// TIA Portal V20 export
// export: Created 2026-10-19T18:06:23.6211165Z, ExportSetting WithDefaults, DisplayName Totally Integrated Automation Portal, DisplayVersion V20 Update 6, DisplayName TIA Portal Openness, DisplayVersion V20 Update 6, DisplayName TIA Portal Version Control Interface, DisplayVersion V20 Update 6, DisplayName SINAMICS Startdrive Advanced, DisplayVersion V20 SP1, DisplayName SINAMICS Startdrive G130, G150, S120, S150, SINAMICS MV, G220, S200, S210, DisplayVersion V20 SP1, DisplayName SINAMICS Startdrive G110M, G120, G120C, G120D, G120P, G115D, DisplayVersion V20 SP1, DisplayName STEP 7 Professional, DisplayVersion V20 Update 6, DisplayName STEP 7 Safety, DisplayVersion V20 Update 2, DisplayName WinCC Basic/Comfort/Advanced, DisplayVersion V20 Update 6, DisplayName WinCC Unified, DisplayVersion V20 Update 6
FUNCTION_BLOCK "SAI_IND_ReadAdjustSettings"   // FB50, LAD
{ S7_Optimized_Access := 'FALSE' }
VERSION : 0.1
// stored: AutoNumber true, IsIECCheckEnabled false, SetENOAutomatically false, UDAEnableTagReadback false
   VAR_INPUT
      ID : HW_IO;   // The Profinet Device Hardware Identifier under device properties
   END_VAR
   VAR_OUTPUT
      ScaleCapacity : Real;   // The configured scale capacity
      Increment : Real;   // The configured scale increment value
      Done : Bool;   // Read done successfully
      Error : Bool;   // Error during reading process
   END_VAR
   VAR_IN_OUT
      Read : Bool;   // Switch this bit ON to start reading
   END_VAR
   VAR DB_SPECIFIC
      Static01 : Bool;
      "Step" : Int;
   END_VAR
   VAR
      RDREC_CAP { S7_SetPoint := 'True'} : RDREC;
   END_VAR
   VAR DB_SPECIFIC
      CAP_RECORD : Real;
      INC_RECORD : Real;
      Activate : Bool;
   END_VAR
   VAR_TEMP
      Temp02 : Bool;
   END_VAR
   VAR_TEMP   // added for the SCL form of the ladder/FBD networks
      _w1 : Bool;
      _w2 : Bool;
      _w3 : Bool;
      _w4 : Bool;
      _w5 : Bool;
      _w6 : Bool;
      _w7 : Bool;
   END_VAR
BEGIN

REGION Network 1: Initialization
   // Initializes FB output bits:
   // Error;
   // Done;
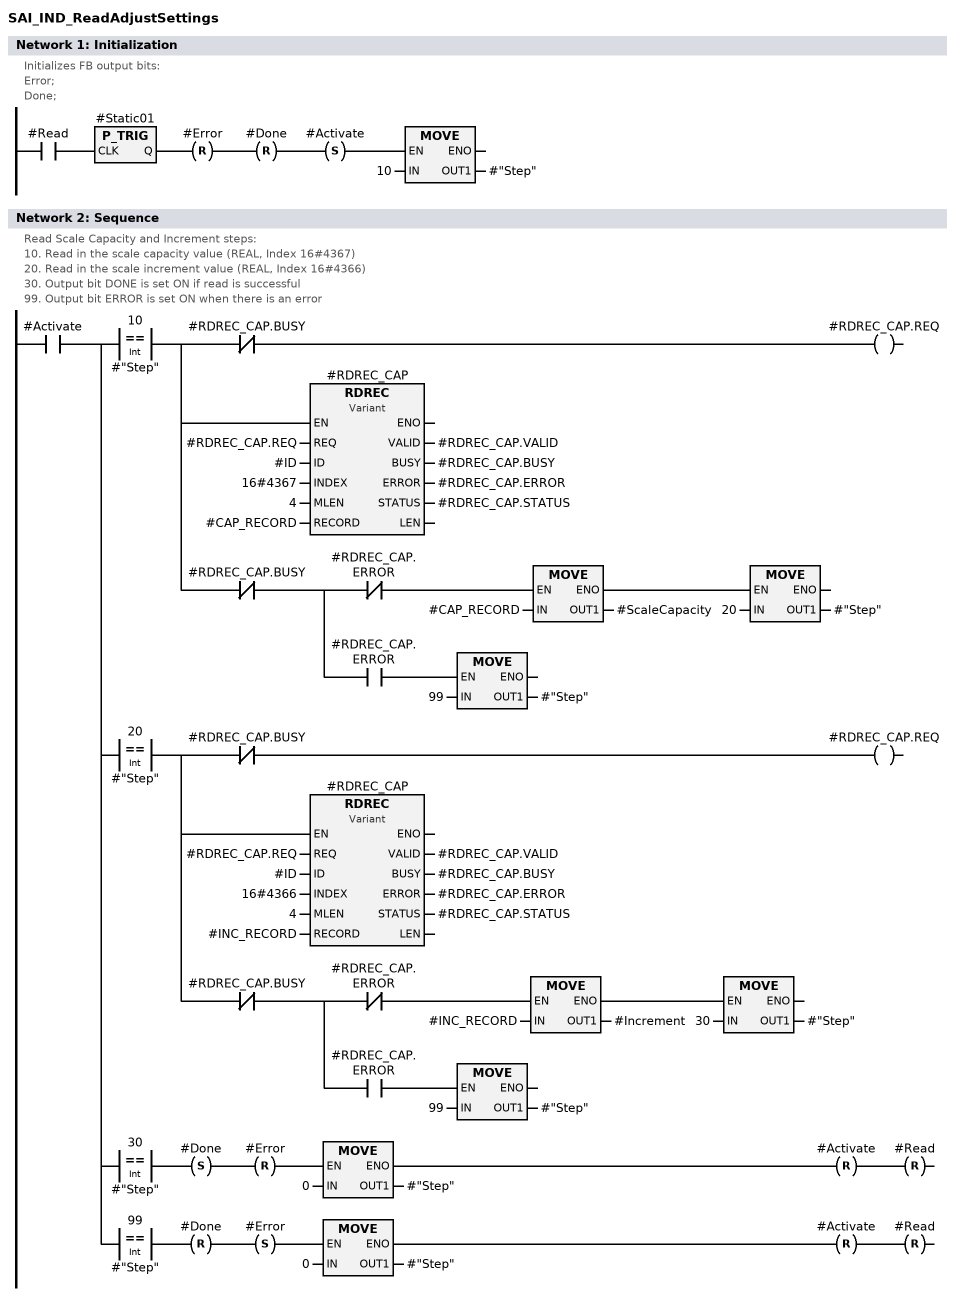
   RUNG wire#powerrail
      Contact( #Read )
      P_Trig( #Static01 )
      R_Coil( #Error )
      R_Coil( #Done )
      S_Coil( #Activate )
      { S7_GenerateENO := "TRUE" } Move(in := 10, out1 => #"Step")
   END_RUNG
   // the same network as SCL:
   #_w1 := #Read AND NOT #Static01;   // rising edge
   #Static01 := #Read;
   IF #_w1 THEN
       #Error := FALSE;
       #Done := FALSE;
       #Activate := TRUE;
       #"Step" := 10;
   END_IF;
END_REGION

REGION Network 2: Sequence
   // Read Scale Capacity and Increment steps:
   // 10. Read in the scale capacity value (REAL, Index 16#4367) 
   // 20. Read in the scale increment value (REAL, Index 16#4366) 
   // 30. Output bit DONE is set ON if read is successful
   // 99. Output bit ERROR is set ON when there is an error
   RUNG wire#powerrail
      Contact( #Activate )
      wire#w1
      { S7_Templates := "SrcType := Int" } EQ_Contact(in1 := 10, in2 := #"Step")
      wire#w2
      I_Contact( #RDREC_CAP.BUSY )
      Coil( #RDREC_CAP.REQ )
   END_RUNG
   RUNG wire#w2
      { S7_Templates := "[ptr_type := Variant, id_type := HW_IO, index_type := DInt, len_type := UInt]" } #RDREC_CAP.RDREC(REQ := #RDREC_CAP.REQ, ID := #ID, INDEX := 16#4367, MLEN := 4, RECORD := #CAP_RECORD, VALID => #RDREC_CAP.VALID, BUSY => #RDREC_CAP.BUSY, ERROR => #RDREC_CAP.ERROR, STATUS => #RDREC_CAP.STATUS, LEN =>)
   END_RUNG
   RUNG wire#w2
      I_Contact( #RDREC_CAP.BUSY )
      wire#w3
      I_Contact( #RDREC_CAP.ERROR )
      { S7_GenerateENO := "TRUE" } Move(in := #CAP_RECORD, out1 => #ScaleCapacity)
      { S7_GenerateENO := "TRUE" } Move(in := 20, out1 => #"Step")
   END_RUNG
   RUNG wire#w3
      Contact( #RDREC_CAP.ERROR )
      { S7_GenerateENO := "TRUE" } Move(in := 99, out1 => #"Step")
   END_RUNG
   RUNG wire#w1
      { S7_Templates := "SrcType := Int" } EQ_Contact(in1 := 20, in2 := #"Step")
      wire#w4
      I_Contact( #RDREC_CAP.BUSY )
      Coil( #RDREC_CAP.REQ )
   END_RUNG
   RUNG wire#w4
      { S7_Templates := "[ptr_type := Variant, id_type := HW_IO, index_type := DInt, len_type := UInt]" } #RDREC_CAP.RDREC(REQ := #RDREC_CAP.REQ, ID := #ID, INDEX := 16#4366, MLEN := 4, RECORD := #INC_RECORD, VALID => #RDREC_CAP.VALID, BUSY => #RDREC_CAP.BUSY, ERROR => #RDREC_CAP.ERROR, STATUS => #RDREC_CAP.STATUS, LEN =>)
   END_RUNG
   RUNG wire#w4
      I_Contact( #RDREC_CAP.BUSY )
      wire#w5
      I_Contact( #RDREC_CAP.ERROR )
      { S7_GenerateENO := "TRUE" } Move(in := #INC_RECORD, out1 => #Increment)
      { S7_GenerateENO := "TRUE" } Move(in := 30, out1 => #"Step")
   END_RUNG
   RUNG wire#w5
      Contact( #RDREC_CAP.ERROR )
      { S7_GenerateENO := "TRUE" } Move(in := 99, out1 => #"Step")
   END_RUNG
   RUNG wire#w1
      { S7_Templates := "SrcType := Int" } EQ_Contact(in1 := 30, in2 := #"Step")
      S_Coil( #Done )
      R_Coil( #Error )
      { S7_GenerateENO := "TRUE" } Move(in := 0, out1 => #"Step")
      R_Coil( #Activate )
      R_Coil( #Read )
   END_RUNG
   RUNG wire#w1
      { S7_Templates := "SrcType := Int" } EQ_Contact(in1 := 99, in2 := #"Step")
      R_Coil( #Done )
      S_Coil( #Error )
      { S7_GenerateENO := "TRUE" } Move(in := 0, out1 => #"Step")
      R_Coil( #Activate )
      R_Coil( #Read )
   END_RUNG
   // the same network as SCL:
   // ENO of a box is taken as its EN; it also drops when the box reports an error
   #_w1 := #Activate AND (10 = #"Step");
   #RDREC_CAP.REQ := #_w1 AND NOT #RDREC_CAP.BUSY;
   IF #_w1 THEN
       #RDREC_CAP(REQ := #RDREC_CAP.REQ,   // RDREC
                  ID := #ID,
                  INDEX := 16#4367,
                  MLEN := 4,
                  RECORD := #CAP_RECORD,
                  VALID => #RDREC_CAP.VALID,
                  BUSY => #RDREC_CAP.BUSY,
                  ERROR => #RDREC_CAP.ERROR,
                  STATUS => #RDREC_CAP.STATUS);
   END_IF;
   #_w2 := #_w1 AND NOT #RDREC_CAP.BUSY;
   IF #_w2 AND NOT #RDREC_CAP.ERROR THEN
       #ScaleCapacity := #CAP_RECORD;
       #"Step" := 20;
   END_IF;
   IF #_w2 AND #RDREC_CAP.ERROR THEN #"Step" := 99; END_IF;
   #_w3 := #Activate AND (20 = #"Step");
   #RDREC_CAP.REQ := #_w3 AND NOT #RDREC_CAP.BUSY;
   IF #_w3 THEN
       #RDREC_CAP(REQ := #RDREC_CAP.REQ,   // RDREC
                  ID := #ID,
                  INDEX := 16#4366,
                  MLEN := 4,
                  RECORD := #INC_RECORD,
                  VALID => #RDREC_CAP.VALID,
                  BUSY => #RDREC_CAP.BUSY,
                  ERROR => #RDREC_CAP.ERROR,
                  STATUS => #RDREC_CAP.STATUS);
   END_IF;
   #_w4 := #_w3 AND NOT #RDREC_CAP.BUSY;
   IF #_w4 AND NOT #RDREC_CAP.ERROR THEN
       #Increment := #INC_RECORD;
       #"Step" := 30;
   END_IF;
   IF #_w4 AND #RDREC_CAP.ERROR THEN #"Step" := 99; END_IF;
   IF #Activate AND (30 = #"Step") THEN
       #Done := TRUE;
       #Error := FALSE;
   END_IF;
   #_w5 := #Activate AND (30 = #"Step");
   IF #_w5 THEN #"Step" := 0; END_IF;
   #_w6 := #Activate;
   IF #_w5 THEN
       #Activate := FALSE;
       #Read := FALSE;
   END_IF;
   IF #_w6 AND (99 = #"Step") THEN
       #Done := FALSE;
       #Error := TRUE;
   END_IF;
   #_w7 := #_w6 AND (99 = #"Step");
   IF #_w7 THEN
       #"Step" := 0;
       #Activate := FALSE;
       #Read := FALSE;
   END_IF;
END_REGION
END_FUNCTION_BLOCK
